TYPE "ST_DeclarationOutImm"
VERSION : 0.1
   STRUCT
      "Sample" : DInt;
   END_STRUCT;
END_TYPE
